Staubli VAL3: logMoveMsgL.pgx

program logMoveMsgL(pointRx x_pPoint, tool x_tTool, mdesc x_mSpeed, num x_nMoveId, bool x_bExact)
  local string l_sCode
  local jointRx l_jRef
  local jointRx l_jResult
  local bool l_bResult
begin
  //
  // 走直线or圆弧时，记录目标点位的joint值参考前一个点的joint（如果是第一次记录，参考herej()）
  if nRecIndex<200
    // l
    if nRecIndex>=1
      l_jRef=jPointRec[nRecIndex-1,1]
    else
      l_jRef=herej()
    endIf
    l_bResult=pointToJoint(x_tTool,l_jRef,x_pPoint,l_jResult)
    //
    if l_bResult==true
      setMutex(bPushToStack)
      jPointRec[nRecIndex,1]=l_jResult
      trToolRec[nRecIndex]=x_tTool.trsf
      mSpeedRec[nRecIndex]=x_mSpeed
      nMoveIdRec[nRecIndex]=x_nMoveId
      bExact[nRecIndex]=x_bExact
      nMoveTypeRec[nRecIndex]=1
      //logMsg("record moveL."+toString("",nMoveIdRec[nRecIndex]))
      nRecIndex=nRecIndex+1
      bPushToStack=false
    else
      // 该位置无关节解
    endIf
  else
    //popUpMsg("记录点数超过容量.")
  endIf

end
